// TIA Portal project "AT3_Start_Uebung" (V18)

(* hardware
DEVICE "PLC_1_Station"  S7-1500 station
   slot 0: "Profilschiene_0"  Rack  6ES7 590-1***0-0AA0
   slot 1: "PLC_1"  CPU 1516-3 PN/DP  6ES7 516-3AN02-0AB0  V2.8
      slot 3: "CPU-Display_1"  6ES7591-1BA00-0AA0
      slot 32768: "PROFINET-Schnittstelle_1"  X1
         slot 32769: "Port_1"  X1 P1
         slot 32770: "Port_2"  X1 P2
      slot 33024: "PROFINET-Schnittstelle_2"  X2
         slot 33025: "Port_1"  X2 P1
      slot 33280: "DP-Schnittstelle_1"  X3
      slot 34817: "Virtual CP interface port_1"  Virtual CP interface port  Virtual CP interface port
   slot 2: "DI_32_HF"  DI 32x24VDC HF  6ES7 521-1BL00-0AB0  V2.2
   slot 3: "DQ_32_ST"  DQ 32x24VDC/0.5A ST  6ES7 522-1BL00-0AB0  V2.0
   slot 4: "AI_8_ST"  AI 8xU/I/RTD/TC ST  6ES7 531-7KF00-0AB0  V2.2
   slot 5: "AQ_4_ST"  AQ 4xU/I ST  6ES7 532-5HD00-0AB0  V2.2
*)

// ===== PLC "PLC_1"  CPU 1516-3 PN/DP =====

VAR_GLOBAL   // PLC tag table "AT3_Grundsteuerung"
   "MotorRechts" AT %Q0.1 : Bool;   // Aus gesicherter Referenz; keine ursprüngliche Laboradresse behauptet.
   "MotorLinks" AT %Q0.2 : Bool;   // Aus gesicherter Referenz; keine ursprüngliche Laboradresse behauptet.
   "SensorLeftHigh" AT %I0.0 : Bool;   // Aus gesicherter Referenz; keine ursprüngliche Laboradresse behauptet.
   "OpticalHigh" AT %I0.1 : Bool;   // Aus gesicherter Referenz; keine ursprüngliche Laboradresse behauptet.
   "SensorRightHigh" AT %I0.2 : Bool;   // Aus gesicherter Referenz; keine ursprüngliche Laboradresse behauptet.
   "HallHigh" AT %I0.3 : Bool;   // Aus gesicherter Referenz; keine ursprüngliche Laboradresse behauptet.
   "LampGreen" AT %Q0.0 : Bool;   // Aus gesicherter Referenz; keine ursprüngliche Laboradresse behauptet.
   "AutomatischeTestMessungAktiv" AT %M0.1 : Bool;   // Aus gesicherter Referenz; keine ursprüngliche Laboradresse behauptet.
   "MessungStartImpuls" AT %M0.3 : Bool;   // Aus gesicherter Referenz; keine ursprüngliche Laboradresse behauptet.
   "LampYellow" AT %Q0.3 : Bool;   // Aus gesicherter Referenz; keine ursprüngliche Laboradresse behauptet.
   "LampRed" AT %Q0.4 : Bool;   // Aus gesicherter Referenz; keine ursprüngliche Laboradresse behauptet.
END_VAR

DATA_BLOCK "HallFlankenZaehler_DB"   // DB2
{ S7_Optimized_Access := 'TRUE' }
AUTHOR : Simatic
FAMILY : IEC
NAME : CNTR
VERSION : 1.0
// stored: InstanceOfName IEC_COUNTER
"IEC_COUNTER"
BEGIN
END_DATA_BLOCK

DATA_BLOCK "Messwerte_DB"   // DB3
{ S7_Optimized_Access := 'TRUE' }
VERSION : 0.1
   VAR
      HallImpulse : Int;   // Aktueller Zählerstand
      MillimeterProImpuls : LReal := 1.2;   // Kalibrierfaktor
      StreckeMm : LReal;   // Berechnete Strecke
      MessungGueltig : Bool;   // TRUE erst nach vollständigem Messzyklus; FALSE bei Zwischenwert oder Abbruch.
   END_VAR
BEGIN
END_DATA_BLOCK

DATA_BLOCK "Motorsteuerung_DB"   // DB4
{ S7_Optimized_Access := 'TRUE' }
VERSION : 0.1
// stored: InstanceOfName Motorsteuerung
"Motorsteuerung"
BEGIN
END_DATA_BLOCK

DATA_BLOCK "Messzyklus_DB"   // DB10
{ S7_Optimized_Access := 'TRUE' }
VERSION : 0.1
// stored: InstanceOfName Messzyklus
"Messzyklus"
BEGIN
END_DATA_BLOCK

DATA_BLOCK "Messauswertung_DB"   // DB11
{ S7_Optimized_Access := 'TRUE' }
VERSION : 0.1
// stored: InstanceOfName Messauswertung
"Messauswertung"
BEGIN
END_DATA_BLOCK

DATA_BLOCK "Ablauf_DB"   // DB12
{ S7_Optimized_Access := 'TRUE' }
// Vorbereitete interne Ablaufmeldungen; keine HMI-Befehle.
   VAR
      HallImpuls : Bool;
      ZyklusBeendet : Bool;
      ZyklusAbgebrochen : Bool;
   END_VAR
BEGIN
END_DATA_BLOCK

FUNCTION_BLOCK "Motorsteuerung"   // FB2, FBD
{ S7_Optimized_Access := 'TRUE' }
VERSION : 0.1
   VAR_INPUT
      RechtsBefehl : Bool;
      LinksBefehl : Bool;
      SensorRechts : Bool;
      SensorLinks : Bool;
      Betriebsfreigabe : Bool;
   END_VAR
   VAR_OUTPUT
      Rechtslauf : Bool;
      Linkslauf : Bool;
   END_VAR
BEGIN

REGION Network 1: Rechtslauf
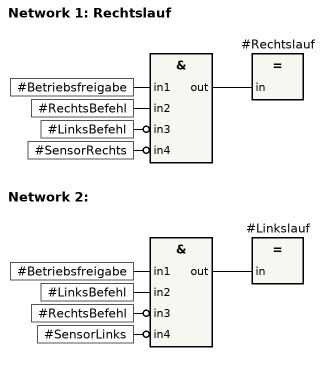
   #Rechtslauf := #Betriebsfreigabe AND #RechtsBefehl AND NOT #LinksBefehl AND NOT #SensorRechts;
END_REGION

REGION Network 2
   #Linkslauf := #Betriebsfreigabe AND #LinksBefehl AND NOT #RechtsBefehl AND NOT #SensorLinks;
END_REGION
END_FUNCTION_BLOCK

FUNCTION_BLOCK "Messzyklus"   // FB10, FBD
{ S7_Optimized_Access := 'TRUE' }
// Rekonstruierter Übungsstart, keine originale Hochschul-Projektdatei.
   VAR_INPUT
      Start : Bool;
      Ende : Bool;
      Abbruch : Bool;
   END_VAR
   VAR_OUTPUT
      Aktiv : Bool;
      Beendet : Bool;
      Abgebrochen : Bool;
   END_VAR
   VAR_TEMP
      VorherAktiv : Bool;
   END_VAR
BEGIN

REGION Network 1: Bisherigen Zustand sichern
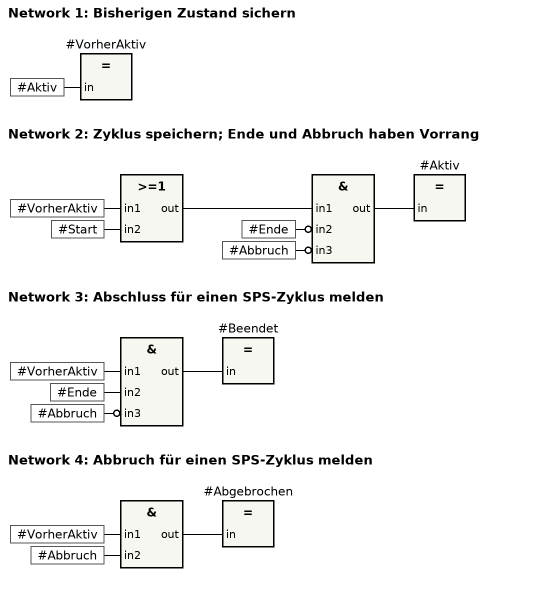
   #VorherAktiv := #Aktiv;
END_REGION

REGION Network 2: Zyklus speichern; Ende und Abbruch haben Vorrang
   // Keine HMI- oder Betriebsartenlogik: Start/Ende/Abbruch kommen ausschließlich aus OB1 Netzwerk 2.
   #Aktiv := (#VorherAktiv OR #Start) AND NOT #Ende AND NOT #Abbruch;
END_REGION

REGION Network 3: Abschluss für einen SPS-Zyklus melden
   #Beendet := #VorherAktiv AND #Ende AND NOT #Abbruch;
END_REGION

REGION Network 4: Abbruch für einen SPS-Zyklus melden
   #Abgebrochen := #VorherAktiv AND #Abbruch;
END_REGION
END_FUNCTION_BLOCK

FUNCTION_BLOCK "Messauswertung"   // FB11, FBD
{ S7_Optimized_Access := 'TRUE' }
// Rekonstruierter Übungsstart, keine originale Hochschul-Projektdatei.
   VAR_INPUT
      ZyklusAktiv : Bool;
      NeuerZyklus : Bool;
      ZyklusEnde : Bool;
      ZyklusAbbruch : Bool;
      Optisch : Bool;
      HallImpuls : Bool;
   END_VAR
   VAR_OUTPUT
      Impulse : Int;
      Gueltig : Bool;
   END_VAR
   VAR
      OptikGesehen : Bool;
      OptikPassiert : Bool;
   END_VAR
BEGIN

REGION Network 1: Echte Hall-Flanken im Messfenster zählen
   // HallImpuls wird ständig vor der Freigabeverknüpfung ermittelt. Stopp ist kein Reset. Nachlaufimpulse werden erfasst, solange der Messzyklus aktiv ist.
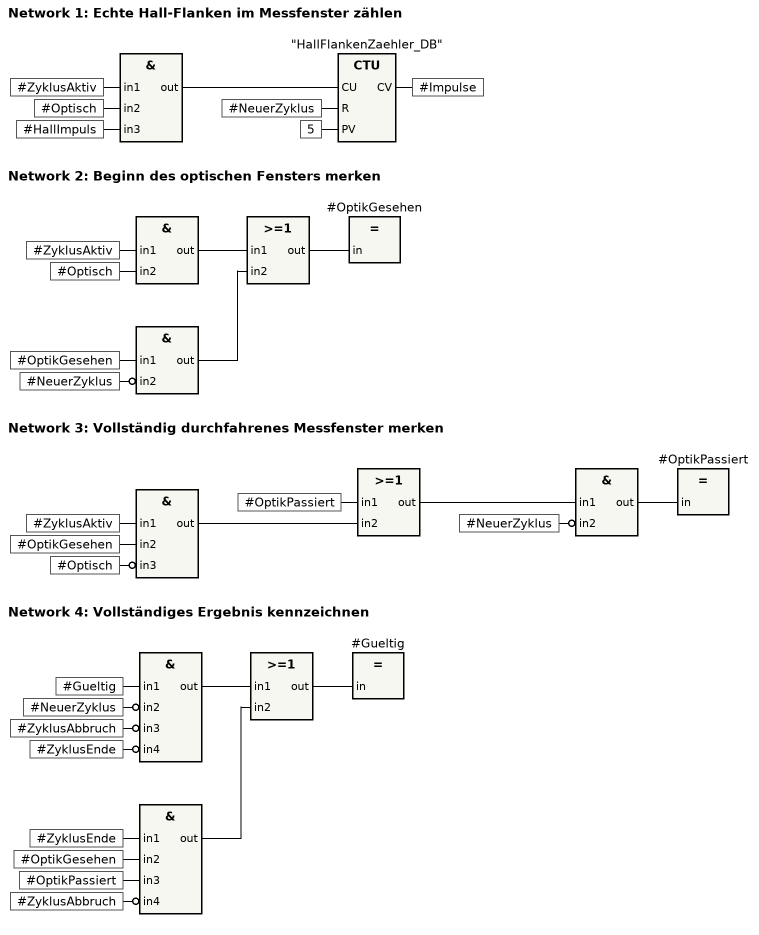
   "HallFlankenZaehler_DB".CTU(CU := #ZyklusAktiv AND #Optisch AND #HallImpuls,
                           R := #NeuerZyklus,
                           PV := 5,
                           CV => #Impulse);
END_REGION

REGION Network 2: Beginn des optischen Fensters merken
   #OptikGesehen := (#ZyklusAktiv AND #Optisch) OR (#OptikGesehen AND NOT #NeuerZyklus);
END_REGION

REGION Network 3: Vollständig durchfahrenes Messfenster merken
   #OptikPassiert := (#OptikPassiert OR (#ZyklusAktiv AND #OptikGesehen AND NOT #Optisch)) AND NOT #NeuerZyklus;
END_REGION

REGION Network 4: Vollständiges Ergebnis kennzeichnen
   // MessungGueltig ist bei neuer oder abgebrochener Messung FALSE; HallImpulse/StreckeMm können dann einen Zwischenwert zeigen.
   #Gueltig := (#Gueltig AND NOT #NeuerZyklus AND NOT #ZyklusAbbruch AND NOT #ZyklusEnde) OR (#ZyklusEnde AND #OptikGesehen AND #OptikPassiert AND NOT #ZyklusAbbruch);
END_REGION
END_FUNCTION_BLOCK

ORGANIZATION_BLOCK "Main"   // OB1, FBD, ProgramCycle
TITLE = "Main Program Sweep (Cycle)"
{ S7_Optimized_Access := 'TRUE' }
VERSION : 0.1
// Rekonstruierter Übungsstart, keine originale Hochschul-Projektdatei.
   VAR_INPUT
      Initial_Call : Bool;   // Initial call of this OB
      Remanence : Bool;   // =True, if remanent data are available
   END_VAR
   VAR_TEMP   // added for the SCL form of the ladder/FBD networks
      _w1 : Bool;
   END_VAR
BEGIN

REGION Network 1: Hall-Flanke erfassen
   // Ständig aufrufen, auch bei stillstehendem Band. Erst die erfasste Flanke wird im Messbaustein mit dem optischen Fenster verknüpft.
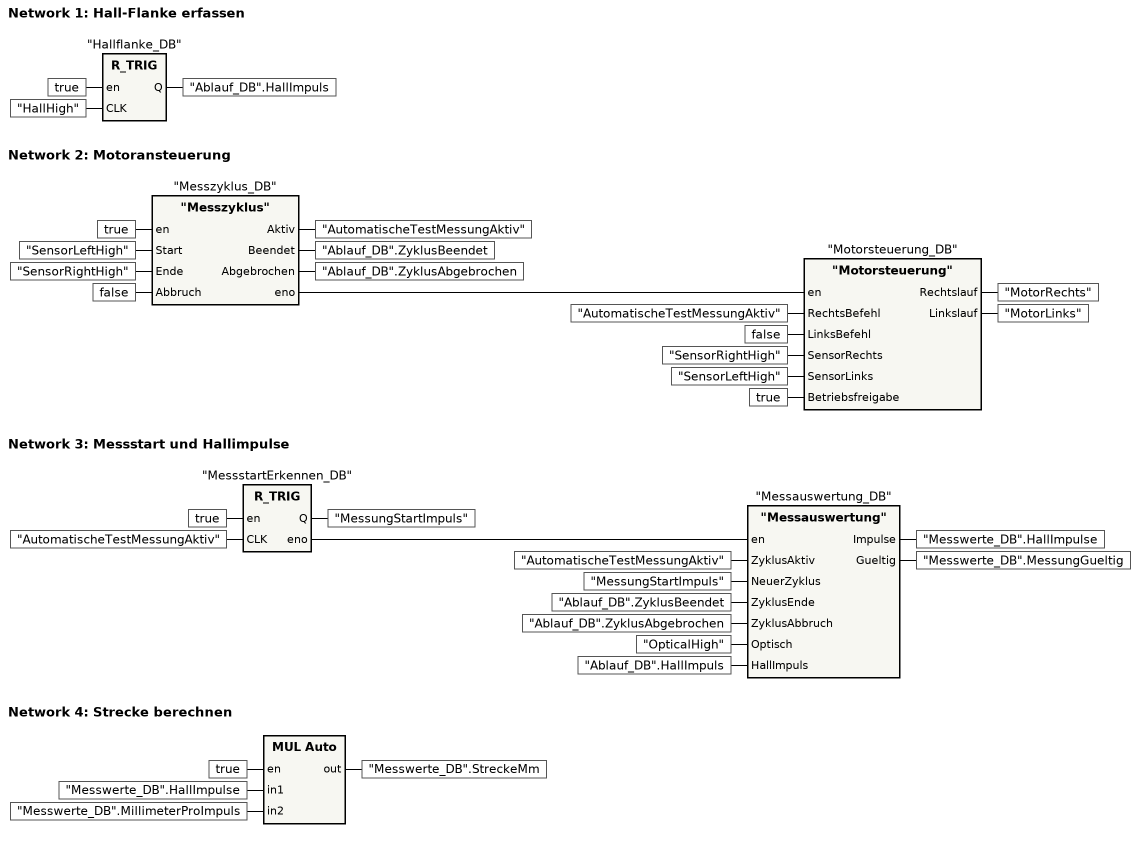
   IF true THEN
       "Hallflanke_DB"(CLK := "HallHigh", Q => "Ablauf_DB".HallImpuls);   // R_TRIG
   END_IF;
END_REGION

REGION Network 2: Motoransteuerung
   // AT-3 Aufgabe 3: Bedienvariablen und ihre Verknüpfungen werden nur hier ergänzt. Stopp sperrt die Betriebsfreigabe, nicht EN; der Zyklus bleibt dabei gespeichert. Messstart/Zählung in Netzwerk 1, 3 und 4 bleiben unverändert.
   "Messzyklus_DB"(EN := true,   // "Messzyklus"
                   Start := "SensorLeftHigh",
                   Ende := "SensorRightHigh",
                   Abbruch := false,
                   Aktiv => "AutomatischeTestMessungAktiv",
                   Beendet => "Ablauf_DB".ZyklusBeendet,
                   Abgebrochen => "Ablauf_DB".ZyklusAbgebrochen,
                   ENO => #_w1);
   IF #_w1 THEN
       "Motorsteuerung_DB"(RechtsBefehl := "AutomatischeTestMessungAktiv",   // "Motorsteuerung"
                           LinksBefehl := false,
                           SensorRechts := "SensorRightHigh",
                           SensorLinks := "SensorLeftHigh",
                           Betriebsfreigabe := true,
                           Rechtslauf => "MotorRechts",
                           Linkslauf => "MotorLinks");
   END_IF;
END_REGION

REGION Network 3: Messstart und Hallimpulse
   // Vorbereitete Messauswertung. Für die Bedienaufgabe nicht ändern. Rücksetzen ausschließlich bei neuem Zyklus; Betriebsstopp setzt nicht zurück.
   // ENO of a box is taken as its EN; it also drops when the box reports an error
   IF true THEN
       "MessstartErkennen_DB"(CLK := "AutomatischeTestMessungAktiv", Q => "MessungStartImpuls");   // R_TRIG
       "Messauswertung_DB"(ZyklusAktiv := "AutomatischeTestMessungAktiv",   // "Messauswertung"
                           NeuerZyklus := "MessungStartImpuls",
                           ZyklusEnde := "Ablauf_DB".ZyklusBeendet,
                           ZyklusAbbruch := "Ablauf_DB".ZyklusAbgebrochen,
                           Optisch := "OpticalHigh",
                           HallImpuls := "Ablauf_DB".HallImpuls,
                           Impulse => "Messwerte_DB".HallImpulse,
                           Gueltig => "Messwerte_DB".MessungGueltig);
   END_IF;
END_REGION

REGION Network 4: Strecke berechnen
   IF true THEN
       "Messwerte_DB".StreckeMm := "Messwerte_DB".HallImpulse * "Messwerte_DB".MillimeterProImpuls;
   END_IF;
END_REGION

REGION Network 5: Ampellogik
   // AT-3 Aufgabe 1.3: Dieses Netzwerk selbst programmieren. Rot: Bandfahrt; Gelb: Längenmessung; Grün: Freigabe für neue Messung.
END_REGION
END_ORGANIZATION_BLOCK